GLOBALCONSTANTS SEC_QUARTER (* Werte einer Section im Condensed Work State (ISO 11783-10), 2 Bit je Section *)
  (* Standard: 61499-2; Description: Copyright (c) 2026 Meisterschulen am Ostbahnhof This program and the accompanying materials are made available under the terms of the Eclipse Public License 2.0 which is available at https://www.eclipse.org/legal/epl-2.0/ SPDX-License-Identifier: EPL-2.0 *)
  (* Version 1.0, 2026-10-31, Franz Höpfinger, Meisterschulen am Ostbahnhof, initial implementation *)
  PACKAGE logiBUS::sections;
  VAR_GLOBAL CONSTANT
    QUARTER_OFF : BYTE := BYTE#2#00; (* aus *)
    QUARTER_ON : BYTE := BYTE#2#01; (* an *)
    QUARTER_ERROR : BYTE := BYTE#2#10; (* Fehler *)
    QUARTER_NA : BYTE := BYTE#2#11; (* nicht verfuegbar *)
  END_VAR
END_GLOBALCONSTANTS
